// SIMATIC S7-200 project (STEP 7-Micro/WIN), CPU 224 CN REL 02.01

SYMBOL_TABLE USUARIO1
SB1R             I1.3     // Pulsador de marcha (verde)
SB2R             I1.2     // Pulsador de paro (rojo)
SA               I1.5     // Selector de modo
QSR              I1.4     // Zeta de emergencia
SM1R             I0.3     // Cilindro largo retraido
SM2R             I0.2     // Cilindro largo extendido
SM3R             I0.1     // Pinza de dedo cerrado
SM4R             I0.4     // Cilindro delgado retraido
SM5R             I0.5     // Cilindro delgado extendido
SF1R             I0.0     // Sensor optico
KB1R             Q0.2     // Accionamiento del cilindro largo
KB2R             Q0.0     // Accionamiento de la pinza
KB3R             Q0.3     // Accionamiento del cilindro delgado
HL1R             Q0.7     // Piloto indicador  de parada
HL2R             Q1.0     // Piloto indicador de marcha
HL3R             Q1.1     // Piloto indicador de emergencia
E0               M0.0     // Estado inicial
E1               M0.1     // Estado para el cierre de la pinza neumatica
E2               M0.2     // Estado para el retroceso del cilindro largo
E3               M0.3     // Estado de salida del cilindro delgado
E4               M0.4     // Estado de retroceso del cilindro delgado
E5               M0.5     // Estado de extension del cilindro largo
E6               M0.6     // Estado de apertura de la garra y avisos
EM               M1.0     // Estado de emergencia
EM1              M1.1     // Estado para la apertura de la garra
EM2              M1.2     // Estado auxiliar para el retorno al estado inicial
EP               M1.3     // Estado de parada
END_SYMBOL_TABLE

ORGANIZATION_BLOCK PRINCIPAL:OB1
TITLE=COMENTARIOS DEL PROGRAMA
BEGIN
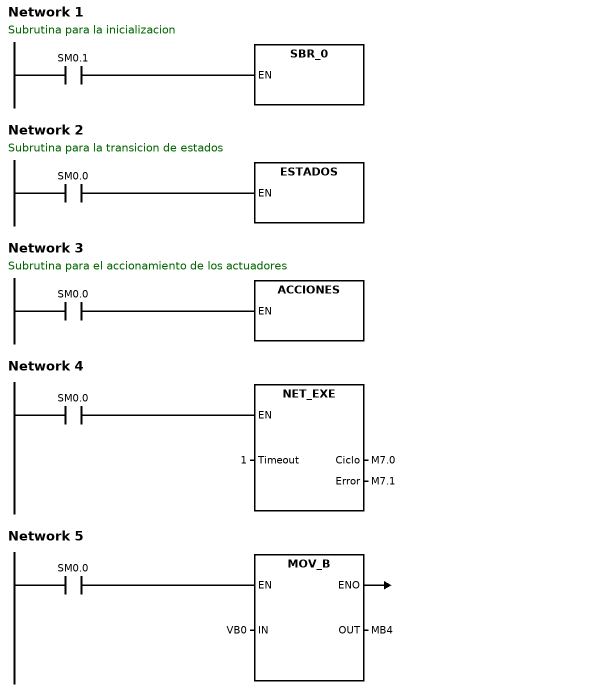
Network 1
// Subrutina para la inicializacion
LD     SM0.1
CALL   SBR_0:SBR0
Network 2
// Subrutina para la transicion de estados
LD     SM0.0
CALL   ESTADOS:SBR1
Network 3
// Subrutina para el accionamiento de los actuadores
LD     SM0.0
CALL   ACCIONES:SBR2
Network 4
LD     SM0.0
CALL   NET_EXE:SBR3, 1, M7.0, M7.1
Network 5
LD     SM0.0
MOVB   VB0, MB4
END_ORGANIZATION_BLOCK

SUBROUTINE_BLOCK SBR_0:SBR0
TITLE=COMENTARIOS DE LA SUBRUTINA
BEGIN
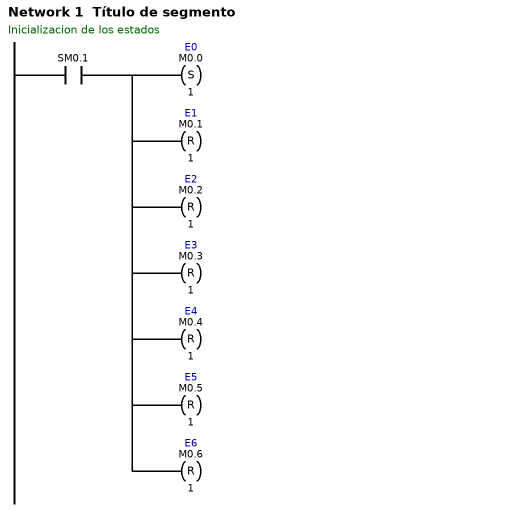
Network 1 // Título de segmento
// Inicializacion de los estados
LD     SM0.1
S      E0:M0.0, 1
R      E1:M0.1, 1
R      E2:M0.2, 1
R      E3:M0.3, 1
R      E4:M0.4, 1
R      E5:M0.5, 1
R      E6:M0.6, 1
END_SUBROUTINE_BLOCK

SUBROUTINE_BLOCK ESTADOS:SBR1
TITLE=TRANSICION DE ESTADOS
BEGIN
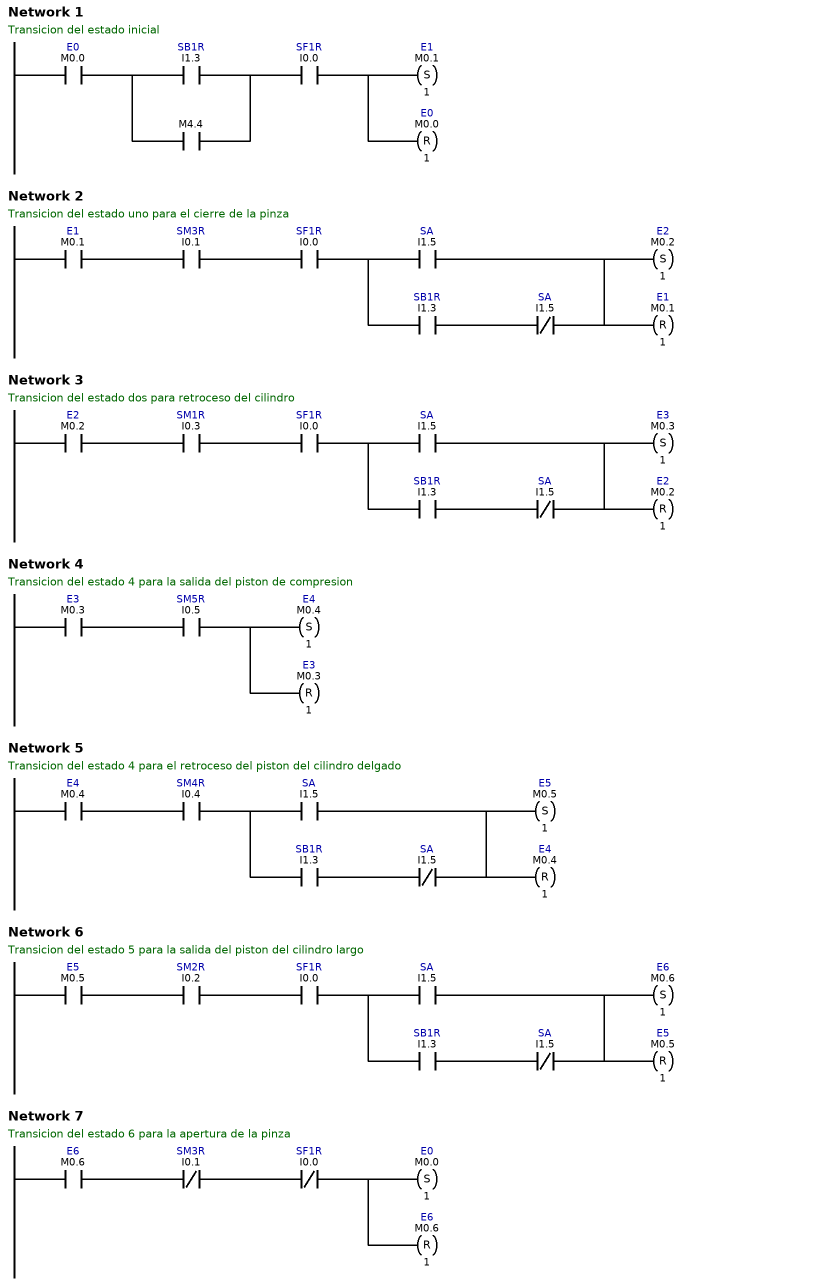
Network 1
// Transicion del estado inicial
LD     E0:M0.0
LD     SB1R:I1.3
O      M4.4
ALD
A      SF1R:I0.0
S      E1:M0.1, 1
R      E0:M0.0, 1
Network 2
// Transicion del estado uno para el cierre de la pinza
LD     E1:M0.1
A      SM3R:I0.1
A      SF1R:I0.0
LD     SA:I1.5
LD     SB1R:I1.3
AN     SA:I1.5
OLD
ALD
S      E2:M0.2, 1
R      E1:M0.1, 1
Network 3
// Transicion del estado dos para retroceso del cilindro
LD     E2:M0.2
A      SM1R:I0.3
A      SF1R:I0.0
LD     SA:I1.5
LD     SB1R:I1.3
AN     SA:I1.5
OLD
ALD
S      E3:M0.3, 1
R      E2:M0.2, 1
Network 4
// Transicion del estado 4 para la salida del piston de compresion
LD     E3:M0.3
A      SM5R:I0.5
S      E4:M0.4, 1
R      E3:M0.3, 1
Network 5
// Transicion del estado 4 para el retroceso del piston del cilindro delgado
LD     E4:M0.4
A      SM4R:I0.4
LD     SA:I1.5
LD     SB1R:I1.3
AN     SA:I1.5
OLD
ALD
S      E5:M0.5, 1
R      E4:M0.4, 1
Network 6
// Transicion del estado 5 para la salida del piston del cilindro largo
LD     E5:M0.5
A      SM2R:I0.2
A      SF1R:I0.0
LD     SA:I1.5
LD     SB1R:I1.3
AN     SA:I1.5
OLD
ALD
S      E6:M0.6, 1
R      E5:M0.5, 1
Network 7
// Transicion del estado 6 para la apertura de la pinza
LD     E6:M0.6
AN     SM3R:I0.1
AN     SF1R:I0.0
S      E0:M0.0, 1
R      E6:M0.6, 1
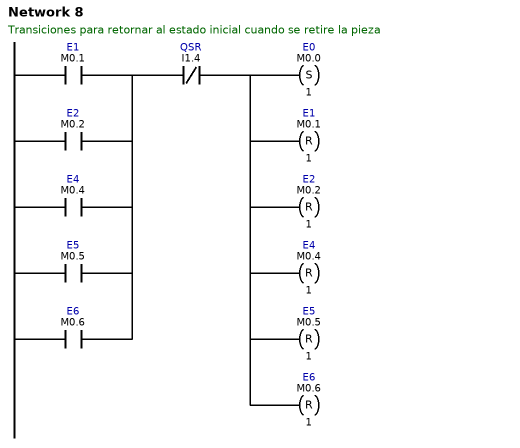
Network 8
// Transiciones para retornar al estado inicial cuando se retire la pieza
LD     E1:M0.1
O      E2:M0.2
O      E4:M0.4
O      E5:M0.5
O      E6:M0.6
AN     QSR:I1.4
S      E0:M0.0, 1
R      E1:M0.1, 1
R      E2:M0.2, 1
R      E4:M0.4, 1
R      E5:M0.5, 1
R      E6:M0.6, 1
END_SUBROUTINE_BLOCK

SUBROUTINE_BLOCK ACCIONES:SBR2
TITLE=SUBRUTINA PARA EL ACCIONAMIENTO DE LOS ACTUADORES
BEGIN
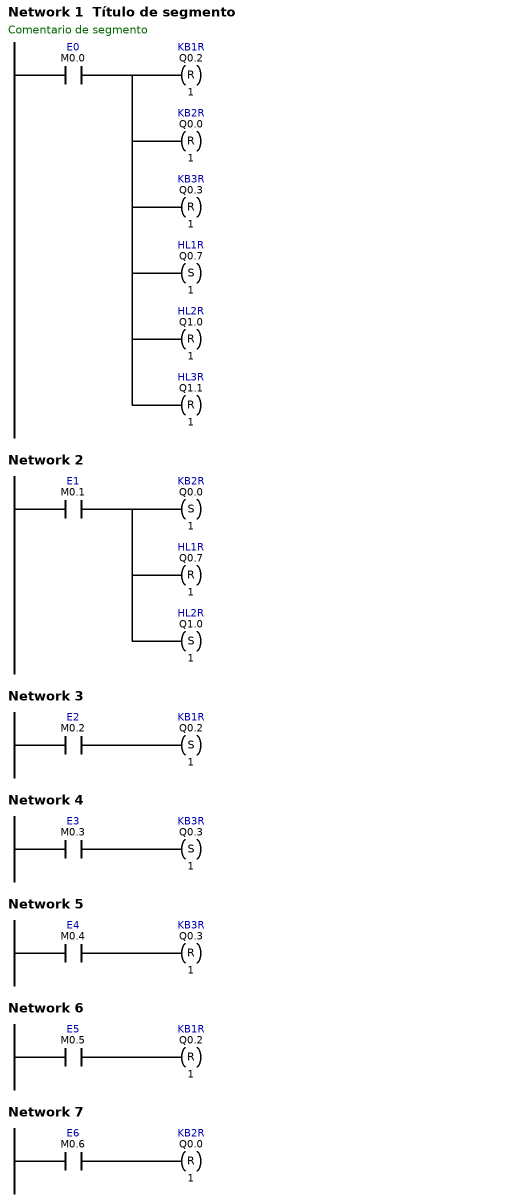
Network 1 // Título de segmento
// Comentario de segmento
LD     E0:M0.0
R      KB1R:Q0.2, 1
R      KB2R:Q0.0, 1
R      KB3R:Q0.3, 1
S      HL1R:Q0.7, 1
R      HL2R:Q1.0, 1
R      HL3R:Q1.1, 1
Network 2
LD     E1:M0.1
S      KB2R:Q0.0, 1
R      HL1R:Q0.7, 1
S      HL2R:Q1.0, 1
Network 3
LD     E2:M0.2
S      KB1R:Q0.2, 1
Network 4
LD     E3:M0.3
S      KB3R:Q0.3, 1
Network 5
LD     E4:M0.4
R      KB3R:Q0.3, 1
Network 6
LD     E5:M0.5
R      KB1R:Q0.2, 1
Network 7
LD     E6:M0.6
R      KB2R:Q0.0, 1
END_SUBROUTINE_BLOCK

// SBR3: protected block, not included
